(* IEC 61131-3 sources: llm-plc-st-eval/data/processed/gpt-4o/B1/zero_shot, 3 files *)

(* ---- ejec_1.st ---- *)
FUNCTION_BLOCK FB_Motor
VAR_INPUT
    btnMarcha : BOOL;   // Botón de marcha
    btnParo : BOOL;     // Botón de paro
    btnEmerg : BOOL;    // Botón de paro de emergencia
END_VAR

VAR_OUTPUT
    motorOn : BOOL;     // Estado del motor
END_VAR

VAR
    motorLatch : BOOL;  // Latch para mantener el estado del motor
    emergStop : BOOL;   // Estado del paro de emergencia
END_VAR

// Inicio del cuerpo del FUNCTION_BLOCK
IF btnEmerg THEN
    // Si el botón de emergencia está presionado, activar el paro de emergencia
    emergStop := TRUE;
    motorLatch := FALSE; // Asegurar que el motor se apague
ELSIF btnParo THEN
    // Si el botón de paro está presionado, apagar el motor
    motorLatch := FALSE;
ELSIF btnMarcha AND NOT emergStop THEN
    // Si el botón de marcha está presionado y no hay paro de emergencia, encender el motor
    motorLatch := TRUE;
END_IF

// Actualizar la salida del motor
motorOn := motorLatch;

// Reiniciar el estado de paro de emergencia si el motor está apagado
IF NOT motorOn THEN
    emergStop := FALSE;
END_IF

END_FUNCTION_BLOCK

(* ---- ejec_2.st ---- *)
FUNCTION_BLOCK FB_Motor
VAR_INPUT
    btnMarcha : BOOL;   // Botón de marcha
    btnParo : BOOL;     // Botón de paro
    btnEmerg : BOOL;    // Botón de paro de emergencia
END_VAR

VAR_OUTPUT
    motorOn : BOOL;     // Estado del motor
END_VAR

VAR
    motorLatch : BOOL;  // Latch para mantener el estado del motor
    emergStopLatch : BOOL; // Latch para mantener el estado de paro de emergencia
END_VAR

// Comportamiento del bloque de función
IF btnEmerg THEN
    // Si el botón de emergencia está presionado, activar el latch de emergencia
    emergStopLatch := TRUE;
    motorLatch := FALSE; // Asegurar que el motor se apague
ELSIF btnParo THEN
    // Si el botón de paro está presionado, apagar el motor
    motorLatch := FALSE;
ELSIF btnMarcha AND NOT emergStopLatch THEN
    // Si el botón de marcha está presionado y no hay paro de emergencia, encender el motor
    motorLatch := TRUE;
END_IF

// Si el paro de emergencia se desactiva, resetear el latch de emergencia
IF NOT btnEmerg THEN
    emergStopLatch := FALSE;
END_IF

// Actualizar la salida del motor
motorOn := motorLatch;

END_FUNCTION_BLOCK

(* ---- ejec_3.st ---- *)
FUNCTION_BLOCK FB_Motor
VAR_INPUT
    btnMarcha : BOOL;   // Botón de marcha
    btnParo   : BOOL;   // Botón de paro
    btnEmerg  : BOOL;   // Botón de paro de emergencia
END_VAR

VAR_OUTPUT
    motorOn   : BOOL;   // Estado del motor (encendido/apagado)
END_VAR

VAR
    motorLatch : BOOL;  // Latch interno para mantener el estado del motor
    emergStopLatch : BOOL; // Latch para el estado de paro de emergencia
END_VAR

// Lógica de control del motor
IF btnEmerg THEN
    // Si se presiona el botón de emergencia, activar el latch de emergencia y apagar el motor
    emergStopLatch := TRUE;
    motorLatch := FALSE;
ELSIF btnParo THEN
    // Si se presiona el botón de paro, apagar el motor
    motorLatch := FALSE;
ELSIF btnMarcha AND NOT emergStopLatch THEN
    // Si se presiona el botón de marcha y no hay paro de emergencia, encender el motor
    motorLatch := TRUE;
END_IF

// El motor está encendido si el latch del motor está activo
motorOn := motorLatch;

// Reset del latch de emergencia si el motor está apagado
IF NOT motorLatch THEN
    emergStopLatch := FALSE;
END_IF

END_FUNCTION_BLOCK
